TYPE ST_AnalogSensor :
STRUCT
	ID		: STRING;
	Value	: REAL;
	Unit	: STRING;
	
	//rawVal_Sensor	: REAL;
	rawVal_Min		: REAL;
	rawVal_Max		: REAL;
	
	outVal_Min		: REAL;
	outVal_Max		: REAL;
	outOffset		: REAL;
	
	//alarms warning
	rLL_Alarm		: REAL	;
	rHH_Alarm		: REAL	;
	rLL_Warning		: REAL	;
	rHH_Warning		: REAL	;
	
END_STRUCT
END_TYPE

(* stored: Version 1.1.0.1, ProductVersion 3.1.4024.12
   DUT ST_AnalogSensor: Id {48421b9c-72bf-4c88-ae11-fcb3ab0e6776} *)
